Fanuc KAREL source: kt00523.KL

-- PROVISIONAL review KL for V770-1; original PC SHA256 7914257a9b955501aa455e16e4ef737cb90f72fe2349e7ab17411281f9894753
-- Incomplete behavior may be omitted. Consult companion uncertainty JSON. Do not deploy.
PROGRAM KT00523
%NOLOCKGROUP
VAR
  OUT : BOOLEAN
-- UNRESOLVED_DECL P1 type=000106
-- UNRESOLVED_DECL P2 type=000106
BEGIN
  -- UNRESOLVED_PC offsets 5-20; opcodes 2E,22,32,35
  -- UNRESOLVED_PC offsets 25-40; opcodes 2E,22,32,35
  -- UNRESOLVED_PC offsets 45-60; opcodes 2E,22,32,35
  -- UNRESOLVED_PC offsets 65-80; opcodes 2E,22,32,35
  -- UNRESOLVED_PC offsets 85-118; opcodes 49,7E,49,7E,AC,23
  -- UNRESOLVED_PC offsets 123-127; opcodes 7F
END KT00523
